(*
SPDX-FileCopyrightText: c 2026 Oleksandr Tiutyk <trofimich@gmail.com>
SPDX-License-Identifier: MIT
License: https://opensource.org/license/mit
*)

(*!
<summary>Checks a direct clone before and after the task-local system wrapper is reconfigured.</summary>
<description>
Uses one task and stays at a stable address while assertions are bound to this instance.
</description>
*)

{attribute 'no_assign'}
{attribute 'no_explicit_call' := 'do not call this function block directly'}
FUNCTION_BLOCK SystemExceptionCloneTest EXTENDS TOF_Testing.SingleCycleTest
VAR_STAT
	{attribute 'hide'}
	_ClassName : STRING := __POUNAME();
END_VAR

(*!
<summary>Checks a direct clone before and after the task-local system wrapper is reconfigured.</summary>
<description>
Supplies native codes to the adapter without raising a native exception. The clone is valid until task cleanup.
</description>
*)
METHOD PROTECTED ExecuteTest
VAR
	original : TOF_Core.IException;
	reconfigured : TOF_Core.IException;
	clonedObject : TOF_Core.IObject;
	cloned : TOF_Core.ISystemException;
	expected : TOF_Core.ERROR_MESSAGE;
	actual : TOF_Core.ERROR_MESSAGE;
	localTimestamp : LDATE_AND_TIME;
	utcTimestamp : LDATE_AND_TIME;
END_VAR
original := TOF_Core.ExceptionManager.GetLastException(
	exceptionCode := __SYSTEM.ExceptionCode.RTSEXCPT_OUT_OF_MEMORY,
	catchPointNamespaceName := 'CloneTest',
	catchPointPOUName := 'OriginalCatch',
	catchPointPosition := 'P1'
);

IF original = 0 THEN
	RecordFailure(message := "The native code must produce a shared wrapper");
	RETURN;
END_IF

expected := original.GetMessage();
localTimestamp := original.LocalTimestamp;
utcTimestamp := original.UtcTimestamp;
clonedObject := original.Clone();

IF NOT __QUERYINTERFACE(clonedObject, cloned) THEN
	RecordFailure(message := "A SystemException clone must implement ISystemException");
	RETURN;
END_IF

Assert.ThatBool(
	actual := cloned.IsDynamicInstance AND_THEN cloned.SelfAddress <> original.SelfAddress,
	message := "The clone must be a distinct task-managed instance"
).IsTrue();

reconfigured := TOF_Core.ExceptionManager.GetLastException(
	exceptionCode := __SYSTEM.ExceptionCode.RTSEXCPT_NOEXCEPTION,
	catchPointNamespaceName := 'Changed',
	catchPointPOUName := 'Changed',
	catchPointPosition := 'P2'
);
Assert.ThatBool(
	actual := reconfigured = original AND_THEN original.Empty,
	message := "The same shared wrapper must be empty after reconfiguration"
).IsTrue();
Assert.ThatBool(
	actual := cloned.ExceptionCode = __SYSTEM.ExceptionCode.RTSEXCPT_OUT_OF_MEMORY,
	message := "The clone must retain the captured native code"
).IsTrue();

actual := cloned.GetMessage();
Assert.ThatBool(
	actual := actual = expected AND_THEN Tc2_Standard.WFIND(STR1 := actual, STR2 := "CloneTest.OriginalCatch at P1") > 0,
	message := "The clone must retain the original diagnostic and catch location"
).IsTrue();
Assert.ThatBool(
	actual := cloned.LocalTimestamp = localTimestamp AND_THEN cloned.UtcTimestamp = utcTimestamp,
	message := "The clone must retain both captured timestamps"
).IsTrue();
END_METHOD

//! <summary>Borrows the concrete class name. Callers must not modify it.</summary>
{attribute 'monitoring' := 'call'}
PROPERTY ClassName : REFERENCE TO STRING
GET
ClassName REF= _ClassName;
END_GET
END_PROPERTY

//! <summary>Borrows the compiler-initialized namespace name. Callers must not modify it.</summary>
{attribute 'monitoring' := 'call'}
PROPERTY NamespaceName : REFERENCE TO STRING
GET
NamespaceName REF= CurrentNamespace.Name;
END_GET
END_PROPERTY

//! <summary>Reports the concrete instance size in bytes.</summary>
{attribute 'monitoring' := 'call'}
PROPERTY SelfSize : ULINT
GET
SelfSize := XSIZEOF(THIS^);
END_GET
END_PROPERTY

END_FUNCTION_BLOCK

(* stored: Version 1.1.0.1
   POU SystemExceptionCloneTest: Id {b08a4e83-4da1-4f60-bec4-ee57cfeda7ca}, SpecialFunc None
   Method ExecuteTest: Id {304d1fcd-4720-44e8-be57-2a0a618a80f6}
   Property ClassName: Id {0b49763c-80f1-4b41-823a-395c775a3391}
   Get Get: Id {76cbe67a-df97-4438-ad71-11cd1faaae86}
   Property NamespaceName: Id {593c0e84-e366-402d-85e7-3a468b017115}
   Get Get: Id {8fcd8407-0aa4-4c60-865a-fdcb8541b637}
   Property SelfSize: Id {f6af564f-71dc-455d-a084-cb2d1620d640}
   Get Get: Id {debdc56d-8165-420a-a824-7ae88a086c69} *)
